Fanuc KAREL source: KA00075.KL

PROGRAM KA00075
%NOLOCKGROUP
VAR
  SRC: XYZWPREXT
  DST: BOOLEAN
BEGIN
  SRC.X = 1.0
  DST = SRC
END KA00075
